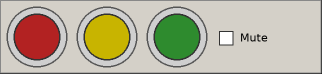
VISUALIZATION Vis_LightTower_1  // 322x74
    Rectangle (0,0 322x74), colour toggle: prg_LightTower.qBuzzer
    Group (2,2 210x70)
        Lamp1 (140,0 70x70), variable: prg_LightTower.qLedGreen, style: Lamp-Lamp1-Green
        Lamp1 (70,0 70x70), variable: prg_LightTower.qLedYellow, style: Lamp-Lamp1-Yellow
        Lamp1 (0,0 70x70), variable: prg_LightTower.qLedRed, style: Lamp-Lamp1-Red
    Checkbox (217,13 95x50), "Mute", variable: bBuzzerMute, input disabled if: prg_User.actUser<2
END_VISUALIZATION

(* stored: Version 1.1.0.1, ProductVersion 3.1.4024.13
   Visu Vis_LightTower_1: Id {c28b9d03-0a4c-47da-b1cc-c49388095387} *)
